// TIA Portal V20 export
// export: Created 2026-10-12T05:42:34.0485366Z, ExportSetting WithDefaults, DisplayName Totally Integrated Automation Portal, DisplayVersion V20, DisplayName TIA Portal Openness, DisplayVersion V20, DisplayName TIA Portal Teamcenter Gateway, DisplayVersion V20, DisplayName TIA Portal Version Control Interface, DisplayVersion V20, DisplayName SINAMICS Startdrive Advanced, DisplayVersion V20 SP1 Update 2, DisplayName SINAMICS Startdrive G110M, G120, G120C, G120D, G120P, G115D, DisplayVersion V20 SP1 Update 2, DisplayName SINAMICS Startdrive G130, G150, S120, S150, SINAMICS MV, G220, S200, S210, DisplayVersion V20 SP1 Update 2, DisplayName STEP 7 Professional, DisplayVersion V20, DisplayName STEP 7 Safety, DisplayVersion V20, DisplayName WinCC Basic/Comfort/Advanced, DisplayVersion V20, DisplayName WinCC Professional, DisplayVersion V20, DisplayName WinCC Unified, DisplayVersion V20
FUNCTION "FRK_CfgRecipe_PressDemoUnit" : Bool   // FC177, SCL
{ S7_Optimized_Access := 'TRUE' }
VERSION : 0.1
// stored: AutoNumber true, IsIECCheckEnabled false, SetENOAutomatically false, UDAEnableTagReadback false
   VAR_INPUT
      ModelCode : String;
      Phase : Int;
   END_VAR
   VAR_IN_OUT
      PressRam : "FB_CylinderCM";
      Door : "FB_CylinderCM";
      PartSlide : "FB_CylinderCM";
      RejectScope : String;
      RejectKey : String;
   END_VAR
   VAR_TEMP
      Ok : Bool;
   END_VAR
BEGIN

   #FRK_CfgRecipe_PressDemoUnit := TRUE;
   #Ok := "FRK_CfgRecipe_CylinderCM"(Module := #PressRam, ModelCode := #ModelCode, Phase := #Phase, RejectScope := #RejectScope, RejectKey := #RejectKey);
   IF NOT #Ok THEN
       #FRK_CfgRecipe_PressDemoUnit := FALSE;
       RETURN;
   END_IF;
   #Ok := "FRK_CfgRecipe_CylinderCM"(Module := #Door, ModelCode := #ModelCode, Phase := #Phase, RejectScope := #RejectScope, RejectKey := #RejectKey);
   IF NOT #Ok THEN
       #FRK_CfgRecipe_PressDemoUnit := FALSE;
       RETURN;
   END_IF;
   #Ok := "FRK_CfgRecipe_CylinderCM"(Module := #PartSlide, ModelCode := #ModelCode, Phase := #Phase, RejectScope := #RejectScope, RejectKey := #RejectKey);
   IF NOT #Ok THEN
       #FRK_CfgRecipe_PressDemoUnit := FALSE;
       RETURN;
   END_IF;
END_FUNCTION
